(* IEC 61131-3 sources: My-first-repository/Branch1_M660.fbsproj/LMC_PacDrive.device.xml.v3^/Plc Logic.plclogic.xml.v3^/Application.application.xml.v3^, 1 file *)

(* ---- SR_Main.prg.st ---- *)
PROGRAM SR_Main
VAR
END_VAR
